FUNCTION_BLOCK SKILL_Run (* One run of a skill primitive, the same for every primitive: waits until the equipment is free, checks the precondition, sends the command, then watches the conditions (or a timer) until the skill is done, has failed or has timed out, and sends the closing command. What the skill is comes in from its contract (SC_). Technical: One run of a skill primitive, the same for every primitive: what the skill is comes in from its contract (socket Contract, AContract); the command goes out to the equipment (plug Equipment, AEquipment) *)
  (* Standard: 61499-2 *)
  (* Version 0.1, 2026-09-28, Project contributors, AAU Smart Production Lab *)
  PACKAGE modlib;
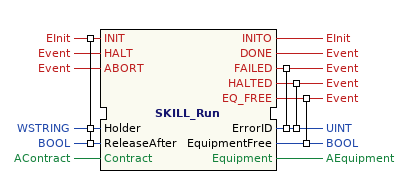
  EVENT_INPUT
    INIT : EInit WITH Holder, ReleaseAfter; (* Initialise: take Holder and ReleaseAfter *)
    HALT; (* Stop the run (ErrorID Interrupted) *)
    ABORT; (* Abort the run: the equipment off and given up *)
  END_EVENT
  EVENT_OUTPUT
    INITO : EInit; (* Initialised: the next block of the INIT chain goes on *)
    DONE; (* The run succeeded *)
    FAILED WITH ErrorID; (* The run failed (ErrorID) *)
    HALTED WITH ErrorID; (* The run was stopped *)
    EQ_FREE WITH EquipmentFree; (* EquipmentFree is updated *)
  END_EVENT
  VAR_INPUT
    Holder : WSTRING; (* The name the equipment is held under: the skill's own, or for a step the skill it belongs to *)
    ReleaseAfter : BOOL; (* Give up the equipment with the run's last command *)
  END_VAR
  VAR_OUTPUT
    ErrorID : UINT; (* Error code: 0 none, 1 PreconditionViolated, 2 InvariantViolated, 3 Timeout, 4 NotReady, 5 NotPermitted, 6 Busy, 7 Interrupted, 8 OutOfRange *)
    EquipmentFree : BOOL; (* The equipment is free, or held under Holder *)
  END_VAR
  SOCKETS
    Contract : modlib::AContract; (* From the skill's contract (AContract): what to do, and when it is done *)
  END_SOCKETS
  PLUGS
    Equipment : modlib::AEquipment; (* To the equipment's port (AEquipment): the commands, PLAYED back *)
  END_PLUGS
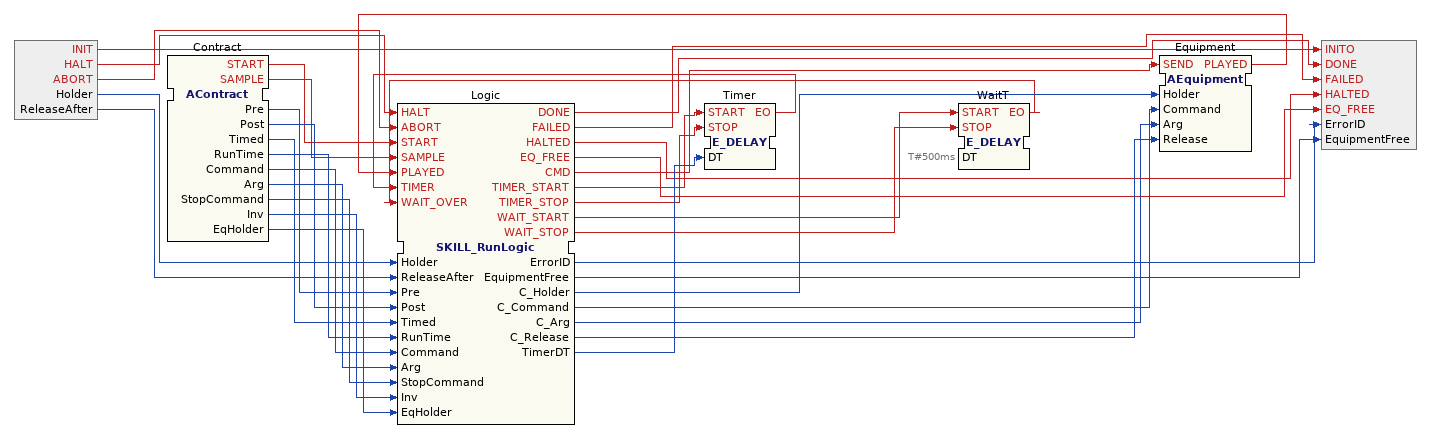
  (* Group OneRun: One run: the contract's values in, the command out, until the end condition or the timer *)
  FBS
    Logic : modlib::SKILL_RunLogic; (* The run's state machine (SKILL_RunLogic). *) {SET_ATTRIBUTE(GroupName, OneRun)}
    Timer : iec61499::events::E_DELAY; (* Ends a skill that runs for a time, or fails a skill that takes longer than its timeout. *) {SET_ATTRIBUTE(GroupName, OneRun)}
    WaitT : iec61499::events::E_DELAY(DT := T#500ms); (* Waits up to half a second for the equipment to become free before giving up (Busy). *) {SET_ATTRIBUTE(GroupName, OneRun)}
  END_FBS
  EVENT_CONNECTIONS
    INIT TO INITO;
    HALT TO Logic.HALT;
    ABORT TO Logic.ABORT;
    Contract.START TO Logic.START;
    Contract.SAMPLE TO Logic.SAMPLE;
    Logic.DONE TO DONE;
    Logic.FAILED TO FAILED;
    Logic.HALTED TO HALTED;
    Logic.EQ_FREE TO EQ_FREE;
    Logic.CMD TO Equipment.SEND;
    Equipment.PLAYED TO Logic.PLAYED;
    Logic.TIMER_START TO Timer.START;
    Logic.TIMER_STOP TO Timer.STOP;
    Timer.EO TO Logic.TIMER;
    Logic.WAIT_START TO WaitT.START;
    Logic.WAIT_STOP TO WaitT.STOP;
    WaitT.EO TO Logic.WAIT_OVER;
  END_CONNECTIONS
  DATA_CONNECTIONS
    Holder TO Logic.Holder;
    ReleaseAfter TO Logic.ReleaseAfter;
    Contract.Pre TO Logic.Pre;
    Contract.Post TO Logic.Post;
    Contract.Timed TO Logic.Timed;
    Contract.RunTime TO Logic.RunTime;
    Contract.Command TO Logic.Command;
    Contract.Arg TO Logic.Arg;
    Contract.StopCommand TO Logic.StopCommand;
    Contract.Inv TO Logic.Inv;
    Contract.EqHolder TO Logic.EqHolder;
    Logic.ErrorID TO ErrorID;
    Logic.EquipmentFree TO EquipmentFree;
    Logic.C_Holder TO Equipment.Holder;
    Logic.C_Command TO Equipment.Command;
    Logic.C_Arg TO Equipment.Arg;
    Logic.C_Release TO Equipment.Release;
    Logic.TimerDT TO Timer.DT;
  END_CONNECTIONS
END_FUNCTION_BLOCK
